(*
SPDX-FileCopyrightText: c 2026 Oleksandr Tiutyk <trofimich@gmail.com>
SPDX-License-Identifier: MIT
License: https://opensource.org/license/mit
*)

(*!
<summary>Groups fixed-capacity queue lookup, FIFO, clear and overflow cases.</summary>
<description>
Owns the independent child instances and their fixed registration array. Use from one PLC task at a stable address.
</description>
*)

{attribute 'no_assign'}
{attribute 'no_explicit_call' := 'do not call this function block directly'}
FUNCTION_BLOCK StaticQueueTestGroup EXTENDS TOF_Testing.TestGroup<6>
VAR_STAT
	{attribute 'hide'}
	_ClassName : STRING := __POUNAME();
END_VAR
VAR
	_Contains : StaticQueueContainsTest(name := "Contains", parent := THIS^);
	_ContainsGeneric : StaticQueueContainsGenericTest(name := "ContainsGeneric", parent := THIS^);
	_EnqueueAndPeek : StaticQueueEnqueueAndPeekTest(name := "EnqueueAndPeek", parent := THIS^);
	_Clear : StaticQueueClearTest(name := "Clear", parent := THIS^);
	_RemoveFirst : StaticQueueRemoveFirstTest(name := "RemoveFirst", parent := THIS^);
	_Overflow : StaticQueueOverflowTest(name := "Overflow", parent := THIS^);

	_Children : ARRAY [0.._ChildCount - 1] OF TOF_Testing.ITestElement :=
	[
		_Contains,
		_ContainsGeneric,
		_EnqueueAndPeek,
		_Clear,
		_RemoveFirst,
		_Overflow
	];
END_VAR

//! <summary>Borrows the fixed child array. Callers must not modify it.</summary>
{attribute 'monitoring' := 'call'}
PROPERTY Children : REFERENCE TO ARRAY [0.._ChildCount - 1] OF TOF_Testing.ITestElement
GET
Children REF= _Children;
END_GET
END_PROPERTY

//! <summary>Borrows the concrete class name. Callers must not modify it.</summary>
{attribute 'monitoring' := 'call'}
PROPERTY ClassName : REFERENCE TO STRING
GET
ClassName REF= _ClassName;
END_GET
END_PROPERTY

//! <summary>Borrows the compiler-initialized namespace name. Callers must not modify it.</summary>
{attribute 'monitoring' := 'call'}
PROPERTY NamespaceName : REFERENCE TO STRING
GET
NamespaceName REF= CurrentNamespace.Name;
END_GET
END_PROPERTY

//! <summary>Reports the concrete instance size in bytes.</summary>
{attribute 'monitoring' := 'call'}
PROPERTY SelfSize : ULINT
GET
SelfSize := XSIZEOF(THIS^);
END_GET
END_PROPERTY

END_FUNCTION_BLOCK

(* stored: Version 1.1.0.1
   POU StaticQueueTestGroup: Id {90d08ca2-ecad-4819-84ab-0582043b3ed0}, SpecialFunc None
   Property Children: Id {5b09ae71-9bba-433a-85d8-437010a6a85e}
   Get Get: Id {285f64ae-7a90-42dd-b9fe-109349f791a3}
   Property ClassName: Id {968580ad-0414-4740-a31c-accdfbe5c78d}
   Get Get: Id {47778292-4dcf-49ee-a6fa-810b02de103d}
   Property NamespaceName: Id {ef516124-c0e0-4901-9a49-37dc2bd124cf}
   Get Get: Id {11c8ed2c-0607-483f-a959-7884e9981670}
   Property SelfSize: Id {31b320c8-fcb0-4fa0-8a88-a770a9c6cdcf}
   Get Get: Id {dc083148-c170-4fe6-a0e3-bb0424b95081} *)
